Fanuc KAREL source: kb00089.KL

-- PROVISIONAL review KL for V770-1; original PC SHA256 fcbe0be7eb35411e3a8df06a52ea158a1b14ef78e2884f18b485d4cab72c55ef
-- Incomplete behavior may be omitted. Consult companion uncertainty JSON. Do not deploy.
PROGRAM KB00089
%NOLOCKGROUP
BEGIN
  -- UNRESOLVED_PC offsets 5-12; opcodes 9D,23
  -- UNRESOLVED_PC offsets 17-24; opcodes 9D,23
  -- UNRESOLVED_PC offsets 29-36; opcodes 9D,23
  -- UNRESOLVED_PC offsets 41-48; opcodes 9D,23
  -- UNRESOLVED_PC offsets 53-60; opcodes 9D,23
  -- UNRESOLVED_PC offsets 65-72; opcodes 9D,23
  -- UNRESOLVED_PC offsets 77-117; opcodes 27,22,22,22,22,22,22,31
  -- UNRESOLVED_PC offsets 122-126; opcodes 7F
END KB00089
